(* Logix 5000 project; controller CIP vendor 1 type 14 code 106 rev 20.12; software revision 20.06; part 12 of 13 *)
(* tags used below, declared in another part *)
   Alarm_Present : INT[8];
   Bit : BOOL[128];
   Counter : COUNTER[10];
   Level_Bits : BOOL[32];
   Level_Timers : TIMER[20];
   MOA_OFF : DINT[10];
   MOA_ON : DINT[10];
   MOA_ONS : DINT;
   MOA_Screen1_Auto : BOOL;
   MOA_Screen1_Man_Off : BOOL;
   MOA_Screen1_Man_On : BOOL;
   MOA_Screen2_Auto : BOOL;
   MOA_Screen2_Man_Off : BOOL;
   MOA_Screen2_Man_On : BOOL;
   MOA_Screen3_Auto : BOOL;
   MOA_Screen3_Man_Off : BOOL;
   MOA_Screen3_Man_On : BOOL;
   MOA_Screen4_Auto : BOOL;
   MOA_Screen4_Man_Off : BOOL;
   MOA_Screen4_Man_On : BOOL;
   MOA_Select : DINT[10];
   MOA_Status : DINT[10];
   MOA_Temp : DINT;
   OpCode_Pin : DINT[5];
   Panelview : INT[40];
   Recipe : RECIPE[41];
   SCLD_Drain_PH : REAL;
   SCLD_Dryer_Duct_Temp : REAL;
   SCLD_Dryer_Exhaust_Temp : REAL;
   SCLD_Return_Temp : REAL;
   SCLD_Rinse_Cond : REAL;
   SCLD_Solution_Tank_Lvl : REAL;
   SCLD_Supply_Temp : REAL;
   SCLD_Wash_Cond : REAL;
   SP_Dryer_Min_Temp : REAL;
   SP_Dryer_Temp : REAL;
   SP_Return_Temp : REAL;
   SP_Rinse_Cond : REAL;
   SP_Solution_Tank_Fill_Lvl : REAL;
   SP_Solution_Tank_Lvl : REAL;
   SP_Supply_Temp : REAL;
   SP_Wash_Cond : REAL;
   SP_Wash_Cond_Hold : REAL;
   Timer : TIMER[99];
   Utility_Out : DINT[5];
   WashChamberDoorGasketCTRL : DINT;
(* MainProgram, continued *)

ROUTINE _30_MAN_OFF_AUTO   (* ladder *)
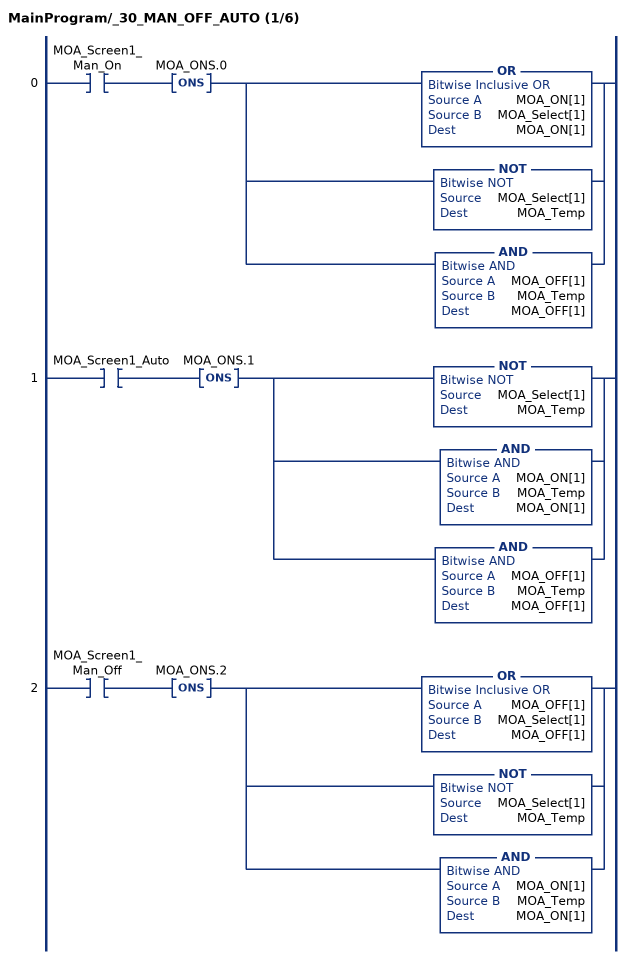
   0: XIC(MOA_Screen1_Man_On)ONS(MOA_ONS.0)[OR(MOA_ON[1],MOA_Select[1],MOA_ON[1]) ,NOT(MOA_Select[1],MOA_Temp) ,AND(MOA_OFF[1],MOA_Temp,MOA_OFF[1]) ];
   1: XIC(MOA_Screen1_Auto)ONS(MOA_ONS.1)[NOT(MOA_Select[1],MOA_Temp) ,AND(MOA_ON[1],MOA_Temp,MOA_ON[1]) ,AND(MOA_OFF[1],MOA_Temp,MOA_OFF[1]) ];
   2: XIC(MOA_Screen1_Man_Off)ONS(MOA_ONS.2)[OR(MOA_OFF[1],MOA_Select[1],MOA_OFF[1]) ,NOT(MOA_Select[1],MOA_Temp) ,AND(MOA_ON[1],MOA_Temp,MOA_ON[1]) ];
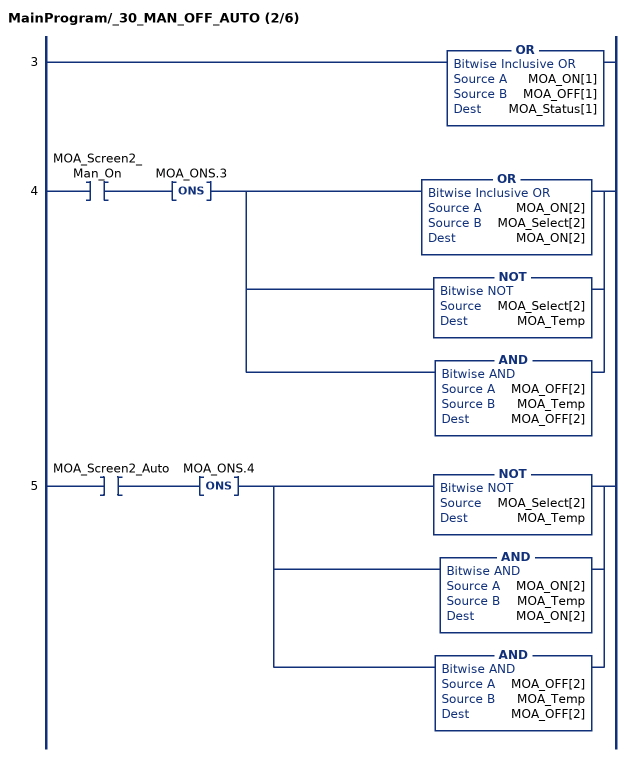
   3: OR(MOA_ON[1],MOA_OFF[1],MOA_Status[1]);
   4: XIC(MOA_Screen2_Man_On)ONS(MOA_ONS.3)[OR(MOA_ON[2],MOA_Select[2],MOA_ON[2]) ,NOT(MOA_Select[2],MOA_Temp) ,AND(MOA_OFF[2],MOA_Temp,MOA_OFF[2]) ];
   5: XIC(MOA_Screen2_Auto)ONS(MOA_ONS.4)[NOT(MOA_Select[2],MOA_Temp) ,AND(MOA_ON[2],MOA_Temp,MOA_ON[2]) ,AND(MOA_OFF[2],MOA_Temp,MOA_OFF[2]) ];
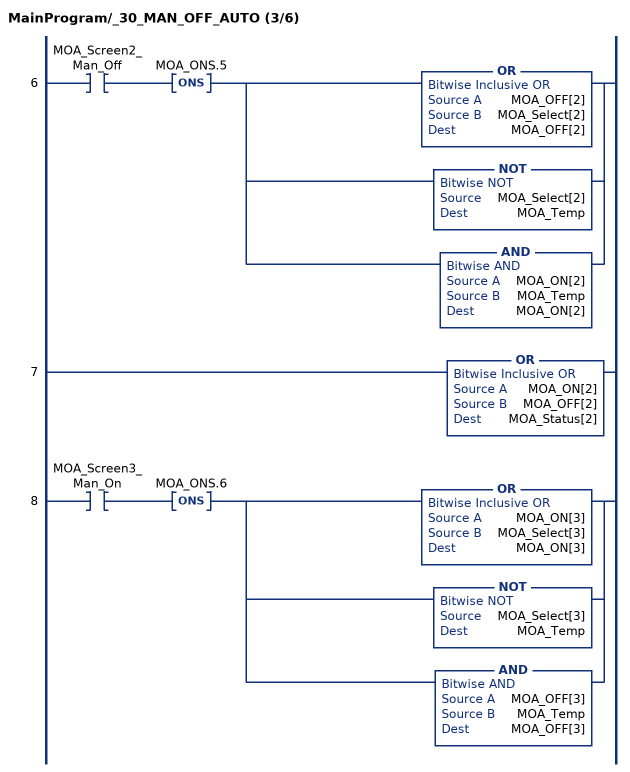
   6: XIC(MOA_Screen2_Man_Off)ONS(MOA_ONS.5)[OR(MOA_OFF[2],MOA_Select[2],MOA_OFF[2]) ,NOT(MOA_Select[2],MOA_Temp) ,AND(MOA_ON[2],MOA_Temp,MOA_ON[2]) ];
   7: OR(MOA_ON[2],MOA_OFF[2],MOA_Status[2]);
   8: XIC(MOA_Screen3_Man_On)ONS(MOA_ONS.6)[OR(MOA_ON[3],MOA_Select[3],MOA_ON[3]) ,NOT(MOA_Select[3],MOA_Temp) ,AND(MOA_OFF[3],MOA_Temp,MOA_OFF[3]) ];
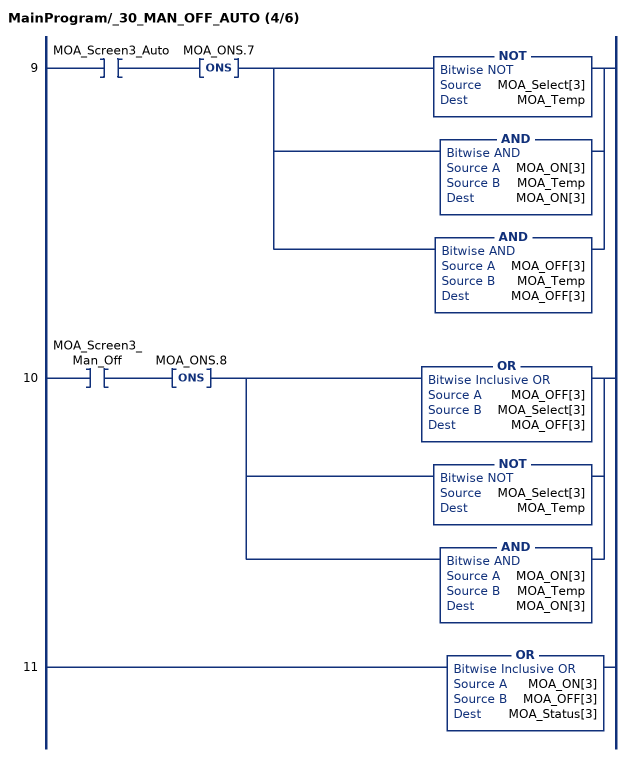
   9: XIC(MOA_Screen3_Auto)ONS(MOA_ONS.7)[NOT(MOA_Select[3],MOA_Temp) ,AND(MOA_ON[3],MOA_Temp,MOA_ON[3]) ,AND(MOA_OFF[3],MOA_Temp,MOA_OFF[3]) ];
   10: XIC(MOA_Screen3_Man_Off)ONS(MOA_ONS.8)[OR(MOA_OFF[3],MOA_Select[3],MOA_OFF[3]) ,NOT(MOA_Select[3],MOA_Temp) ,AND(MOA_ON[3],MOA_Temp,MOA_ON[3]) ];
   11: OR(MOA_ON[3],MOA_OFF[3],MOA_Status[3]);
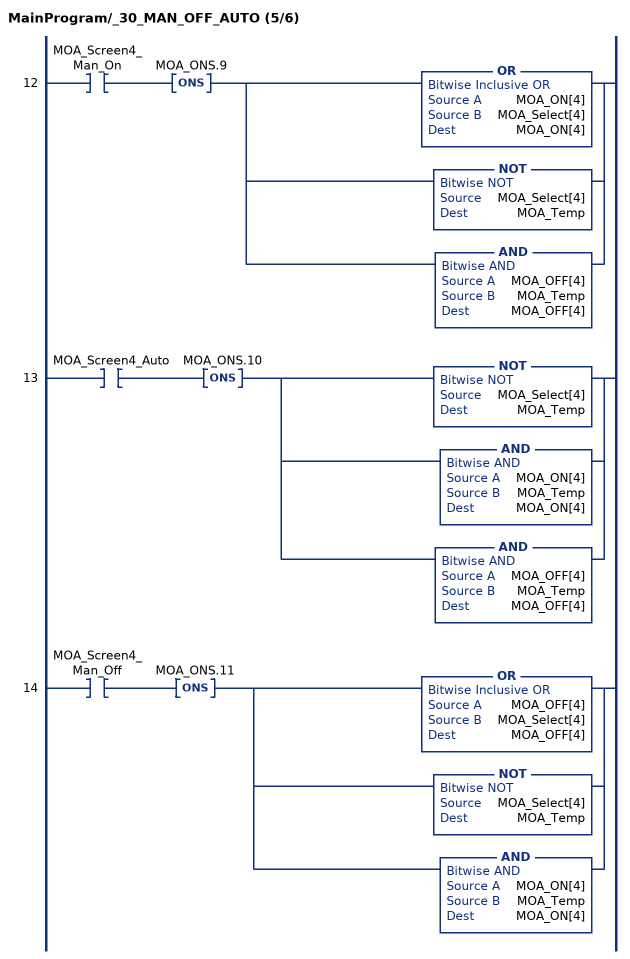
   12: XIC(MOA_Screen4_Man_On)ONS(MOA_ONS.9)[OR(MOA_ON[4],MOA_Select[4],MOA_ON[4]) ,NOT(MOA_Select[4],MOA_Temp) ,AND(MOA_OFF[4],MOA_Temp,MOA_OFF[4]) ];
   13: XIC(MOA_Screen4_Auto)ONS(MOA_ONS.10)[NOT(MOA_Select[4],MOA_Temp) ,AND(MOA_ON[4],MOA_Temp,MOA_ON[4]) ,AND(MOA_OFF[4],MOA_Temp,MOA_OFF[4]) ];
   14: XIC(MOA_Screen4_Man_Off)ONS(MOA_ONS.11)[OR(MOA_OFF[4],MOA_Select[4],MOA_OFF[4]) ,NOT(MOA_Select[4],MOA_Temp) ,AND(MOA_ON[4],MOA_Temp,MOA_ON[4]) ];
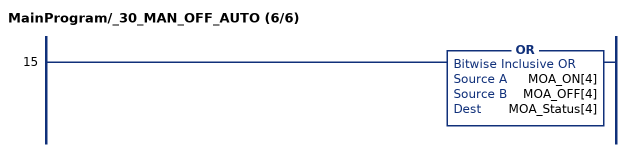
   15: OR(MOA_ON[4],MOA_OFF[4],MOA_Status[4]);
END_ROUTINE

ROUTINE _80_DOOR_GASKET   (* ladder *)
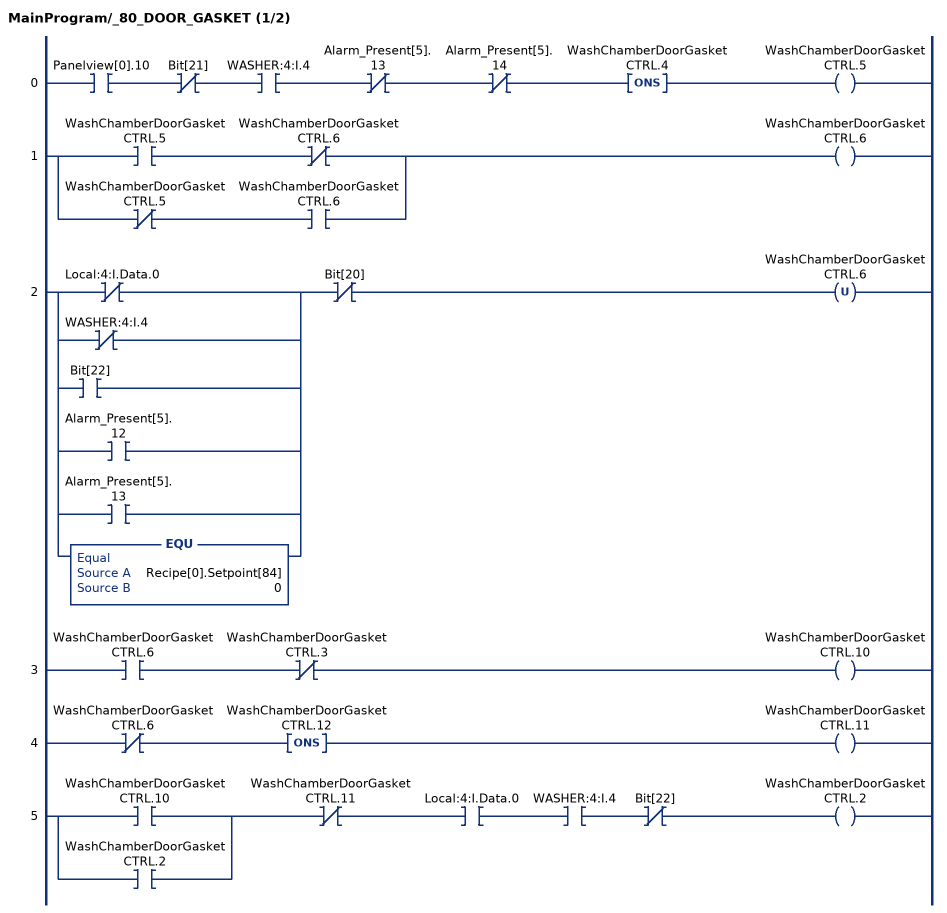
   0: XIC(Panelview[0].10)XIO(Bit[21])XIC(WASHER:4:I.4)XIO(Alarm_Present[5].13)XIO(Alarm_Present[5].14)ONS(WashChamberDoorGasketCTRL.4)OTE(WashChamberDoorGasketCTRL.5);
   1: [XIC(WashChamberDoorGasketCTRL.5) XIO(WashChamberDoorGasketCTRL.6) ,XIO(WashChamberDoorGasketCTRL.5) XIC(WashChamberDoorGasketCTRL.6) ]OTE(WashChamberDoorGasketCTRL.6);
   2: [XIO(Local:4:I.Data.0) ,XIO(WASHER:4:I.4) ,XIC(Bit[22]) ,XIC(Alarm_Present[5].12) ,XIC(Alarm_Present[5].13) ,EQU(Recipe[0].Setpoint[84],0) ]XIO(Bit[20])OTU(WashChamberDoorGasketCTRL.6);
   3: XIC(WashChamberDoorGasketCTRL.6)XIO(WashChamberDoorGasketCTRL.3)OTE(WashChamberDoorGasketCTRL.10);
   4: XIO(WashChamberDoorGasketCTRL.6)ONS(WashChamberDoorGasketCTRL.12)OTE(WashChamberDoorGasketCTRL.11);
   5: [XIC(WashChamberDoorGasketCTRL.10) ,XIC(WashChamberDoorGasketCTRL.2) ]XIO(WashChamberDoorGasketCTRL.11)XIC(Local:4:I.Data.0)XIC(WASHER:4:I.4)XIO(Bit[22])OTE(WashChamberDoorGasketCTRL.2);
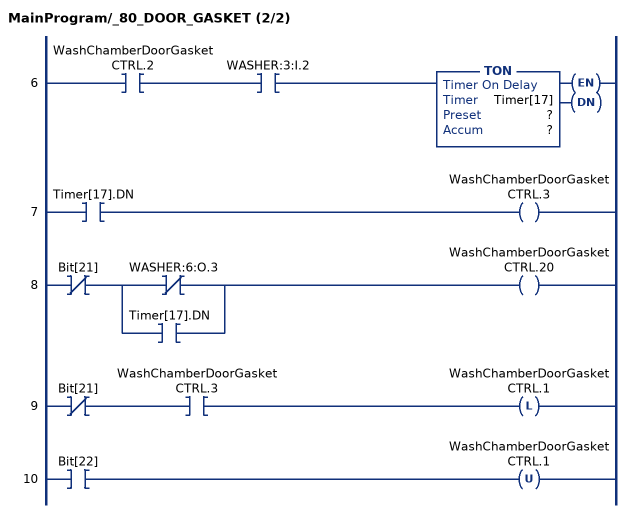
   6: XIC(WashChamberDoorGasketCTRL.2)XIC(WASHER:3:I.2)TON(Timer[17],?,?);
   7: XIC(Timer[17].DN)OTE(WashChamberDoorGasketCTRL.3);
   8: XIO(Bit[21])[XIO(WASHER:6:O.3) ,XIC(Timer[17].DN) ]OTE(WashChamberDoorGasketCTRL.20);
   9: XIO(Bit[21])XIC(WashChamberDoorGasketCTRL.3)OTL(WashChamberDoorGasketCTRL.1);
   10: XIC(Bit[22])OTU(WashChamberDoorGasketCTRL.1);
END_ROUTINE

ROUTINE _86_TEMPERATURE   (* ladder *)
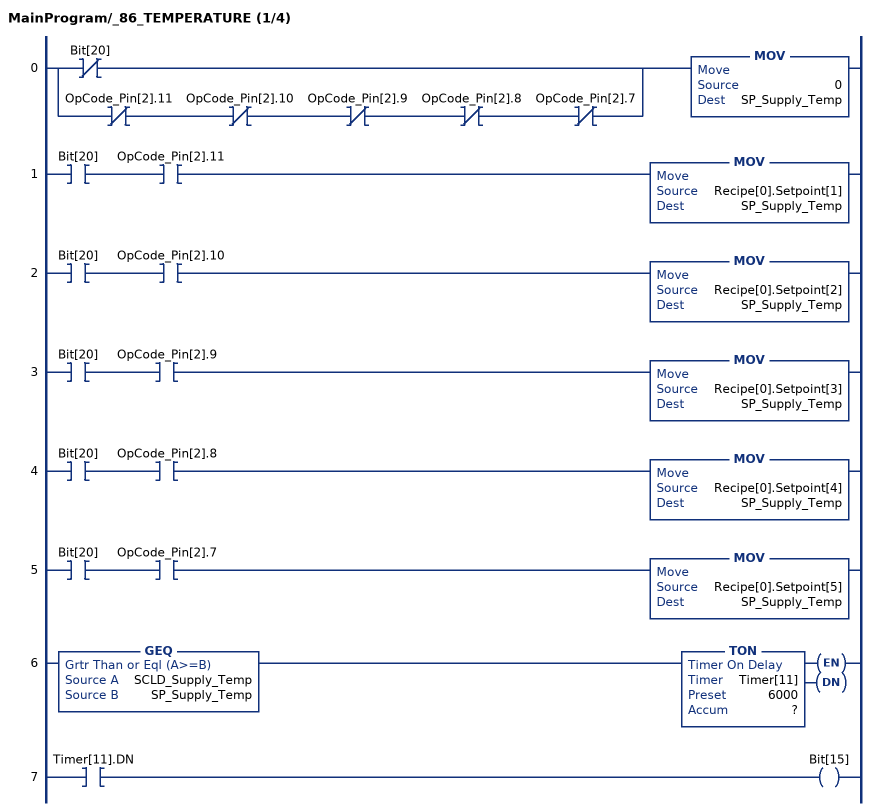
   0: [XIO(Bit[20]) ,XIO(OpCode_Pin[2].11) XIO(OpCode_Pin[2].10) XIO(OpCode_Pin[2].9) XIO(OpCode_Pin[2].8) XIO(OpCode_Pin[2].7) ]MOV(0,SP_Supply_Temp);
   1: XIC(Bit[20])XIC(OpCode_Pin[2].11)MOV(Recipe[0].Setpoint[1],SP_Supply_Temp);
   2: XIC(Bit[20])XIC(OpCode_Pin[2].10)MOV(Recipe[0].Setpoint[2],SP_Supply_Temp);
   3: XIC(Bit[20])XIC(OpCode_Pin[2].9)MOV(Recipe[0].Setpoint[3],SP_Supply_Temp);
   4: XIC(Bit[20])XIC(OpCode_Pin[2].8)MOV(Recipe[0].Setpoint[4],SP_Supply_Temp);
   5: XIC(Bit[20])XIC(OpCode_Pin[2].7)MOV(Recipe[0].Setpoint[5],SP_Supply_Temp);
   6: GEQ(SCLD_Supply_Temp,SP_Supply_Temp)TON(Timer[11],?,?);
   7: XIC(Timer[11].DN)OTE(Bit[15]);
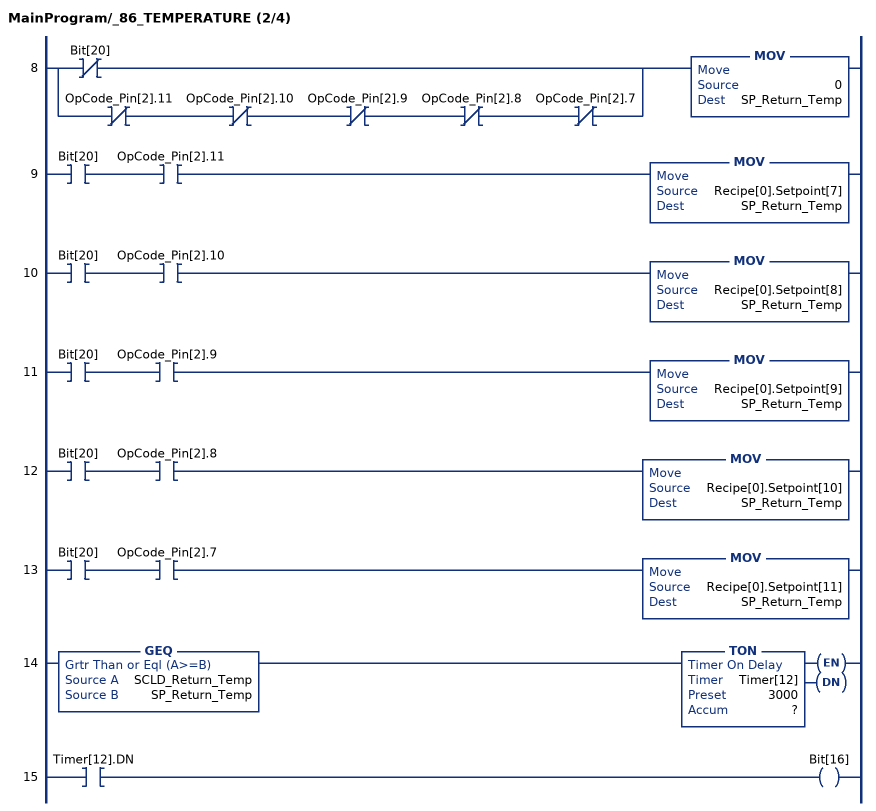
   8: [XIO(Bit[20]) ,XIO(OpCode_Pin[2].11) XIO(OpCode_Pin[2].10) XIO(OpCode_Pin[2].9) XIO(OpCode_Pin[2].8) XIO(OpCode_Pin[2].7) ]MOV(0,SP_Return_Temp);
   9: XIC(Bit[20])XIC(OpCode_Pin[2].11)MOV(Recipe[0].Setpoint[7],SP_Return_Temp);
   10: XIC(Bit[20])XIC(OpCode_Pin[2].10)MOV(Recipe[0].Setpoint[8],SP_Return_Temp);
   11: XIC(Bit[20])XIC(OpCode_Pin[2].9)MOV(Recipe[0].Setpoint[9],SP_Return_Temp);
   12: XIC(Bit[20])XIC(OpCode_Pin[2].8)MOV(Recipe[0].Setpoint[10],SP_Return_Temp);
   13: XIC(Bit[20])XIC(OpCode_Pin[2].7)MOV(Recipe[0].Setpoint[11],SP_Return_Temp);
   14: GEQ(SCLD_Return_Temp,SP_Return_Temp)TON(Timer[12],?,?);
   15: XIC(Timer[12].DN)OTE(Bit[16]);
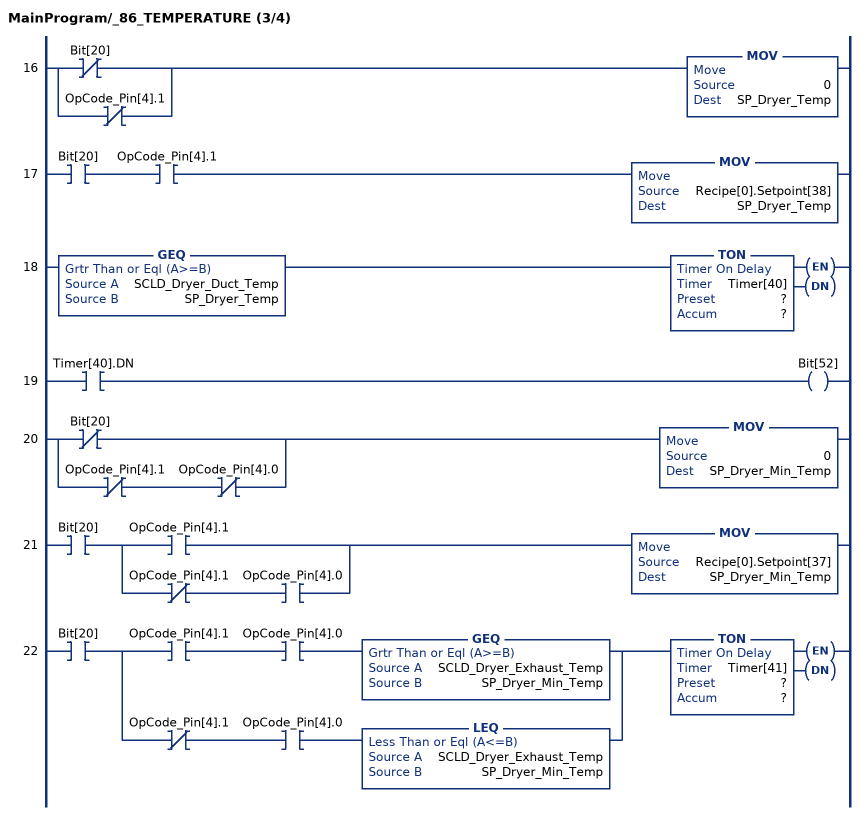
   16: [XIO(Bit[20]) ,XIO(OpCode_Pin[4].1) ]MOV(0,SP_Dryer_Temp);
   17: XIC(Bit[20])XIC(OpCode_Pin[4].1)MOV(Recipe[0].Setpoint[38],SP_Dryer_Temp);
   18: GEQ(SCLD_Dryer_Duct_Temp,SP_Dryer_Temp)TON(Timer[40],?,?);
   19: XIC(Timer[40].DN)OTE(Bit[52]);
   20: [XIO(Bit[20]) ,XIO(OpCode_Pin[4].1) XIO(OpCode_Pin[4].0) ]MOV(0,SP_Dryer_Min_Temp);
   21: XIC(Bit[20])[XIC(OpCode_Pin[4].1) ,XIO(OpCode_Pin[4].1) XIC(OpCode_Pin[4].0) ]MOV(Recipe[0].Setpoint[37],SP_Dryer_Min_Temp);
   22: XIC(Bit[20])[XIC(OpCode_Pin[4].1) XIC(OpCode_Pin[4].0) GEQ(SCLD_Dryer_Exhaust_Temp,SP_Dryer_Min_Temp) ,XIO(OpCode_Pin[4].1) XIC(OpCode_Pin[4].0) LEQ(SCLD_Dryer_Exhaust_Temp,SP_Dryer_Min_Temp) ]TON(Timer[41],?,?);
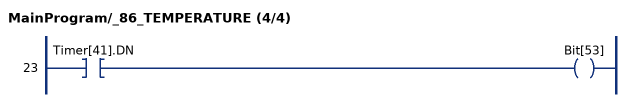
   23: XIC(Timer[41].DN)OTE(Bit[53]);
END_ROUTINE

ROUTINE _87_CONDUCTIVITY   (* ladder *)
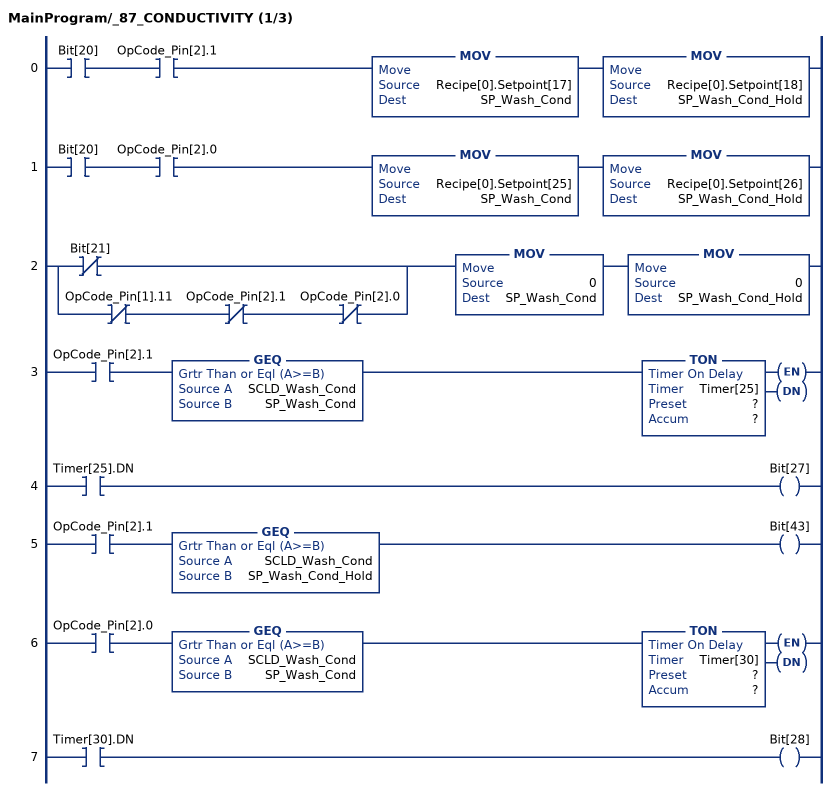
   0: XIC(Bit[20])XIC(OpCode_Pin[2].1)MOV(Recipe[0].Setpoint[17],SP_Wash_Cond)MOV(Recipe[0].Setpoint[18],SP_Wash_Cond_Hold);
   1: XIC(Bit[20])XIC(OpCode_Pin[2].0)MOV(Recipe[0].Setpoint[25],SP_Wash_Cond)MOV(Recipe[0].Setpoint[26],SP_Wash_Cond_Hold);
   2: [XIO(Bit[21]) ,XIO(OpCode_Pin[1].11) XIO(OpCode_Pin[2].1) XIO(OpCode_Pin[2].0) ]MOV(0,SP_Wash_Cond)MOV(0,SP_Wash_Cond_Hold);
   3: XIC(OpCode_Pin[2].1)GEQ(SCLD_Wash_Cond,SP_Wash_Cond)TON(Timer[25],?,?);
   4: XIC(Timer[25].DN)OTE(Bit[27]);
   5: XIC(OpCode_Pin[2].1)GEQ(SCLD_Wash_Cond,SP_Wash_Cond_Hold)OTE(Bit[43]);
   6: XIC(OpCode_Pin[2].0)GEQ(SCLD_Wash_Cond,SP_Wash_Cond)TON(Timer[30],?,?);
   7: XIC(Timer[30].DN)OTE(Bit[28]);
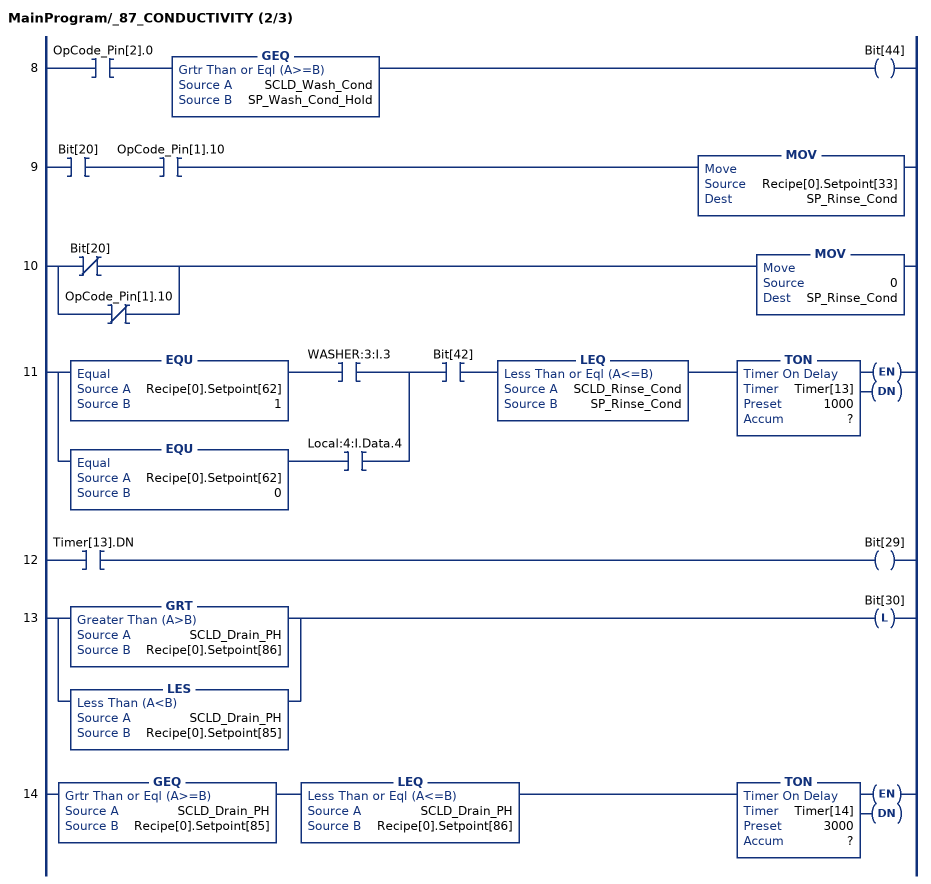
   8: XIC(OpCode_Pin[2].0)GEQ(SCLD_Wash_Cond,SP_Wash_Cond_Hold)OTE(Bit[44]);
   9: XIC(Bit[20])XIC(OpCode_Pin[1].10)MOV(Recipe[0].Setpoint[33],SP_Rinse_Cond);
   10: [XIO(Bit[20]) ,XIO(OpCode_Pin[1].10) ]MOV(0,SP_Rinse_Cond);
   11: [EQU(Recipe[0].Setpoint[62],1) XIC(WASHER:3:I.3) ,EQU(Recipe[0].Setpoint[62],0) XIC(Local:4:I.Data.4) ]XIC(Bit[42])LEQ(SCLD_Rinse_Cond,SP_Rinse_Cond)TON(Timer[13],?,?);
   12: XIC(Timer[13].DN)OTE(Bit[29]);
   13: [GRT(SCLD_Drain_PH,Recipe[0].Setpoint[86]) ,LES(SCLD_Drain_PH,Recipe[0].Setpoint[85]) ]OTL(Bit[30]);
   14: GEQ(SCLD_Drain_PH,Recipe[0].Setpoint[85])LEQ(SCLD_Drain_PH,Recipe[0].Setpoint[86])TON(Timer[14],?,?);
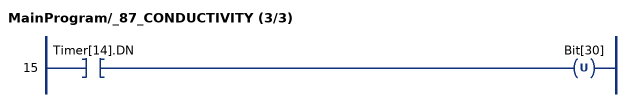
   15: XIC(Timer[14].DN)OTU(Bit[30]);
END_ROUTINE

ROUTINE _88_LEVEL   (* ladder *)
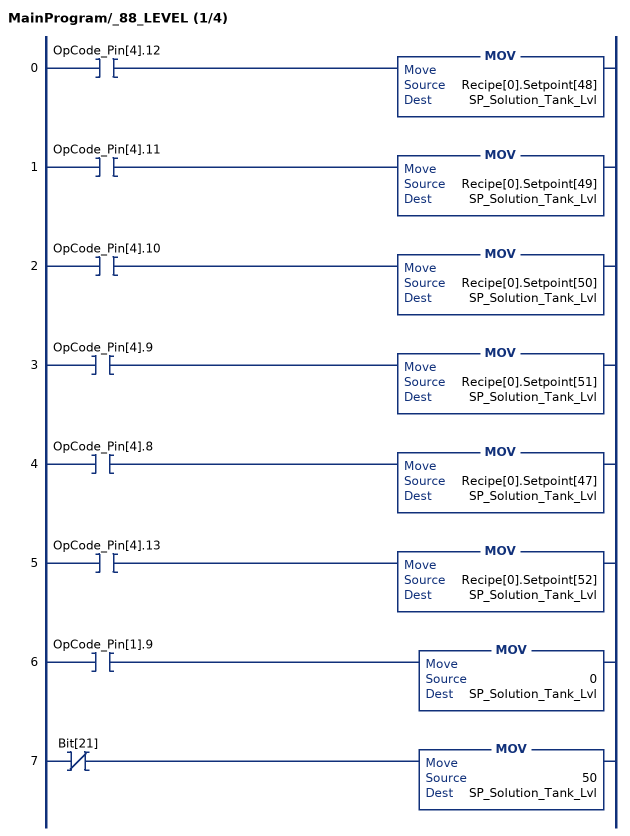
   0: XIC(OpCode_Pin[4].12)MOV(Recipe[0].Setpoint[48],SP_Solution_Tank_Lvl);
   1: XIC(OpCode_Pin[4].11)MOV(Recipe[0].Setpoint[49],SP_Solution_Tank_Lvl);
   2: XIC(OpCode_Pin[4].10)MOV(Recipe[0].Setpoint[50],SP_Solution_Tank_Lvl);
   3: XIC(OpCode_Pin[4].9)MOV(Recipe[0].Setpoint[51],SP_Solution_Tank_Lvl);
   4: XIC(OpCode_Pin[4].8)MOV(Recipe[0].Setpoint[47],SP_Solution_Tank_Lvl);
   5: XIC(OpCode_Pin[4].13)MOV(Recipe[0].Setpoint[52],SP_Solution_Tank_Lvl);
   6: XIC(OpCode_Pin[1].9)MOV(0,SP_Solution_Tank_Lvl);
   7: XIO(Bit[21])MOV(50,SP_Solution_Tank_Lvl);
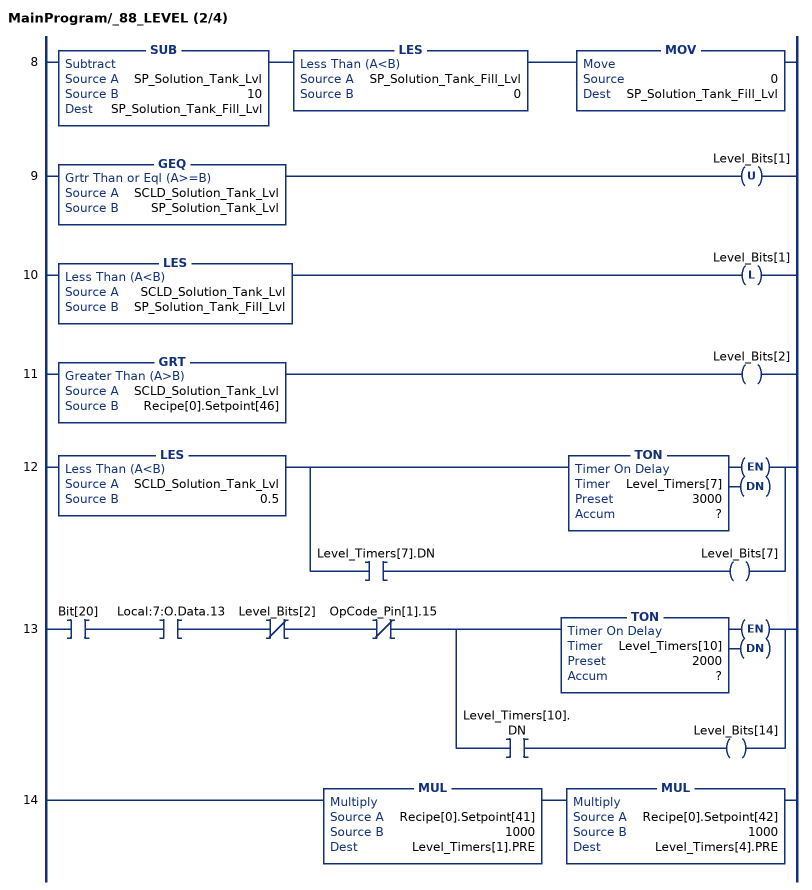
   8: SUB(SP_Solution_Tank_Lvl,10,SP_Solution_Tank_Fill_Lvl)LES(SP_Solution_Tank_Fill_Lvl,0)MOV(0,SP_Solution_Tank_Fill_Lvl);
   9: GEQ(SCLD_Solution_Tank_Lvl,SP_Solution_Tank_Lvl)OTU(Level_Bits[1]);
   10: LES(SCLD_Solution_Tank_Lvl,SP_Solution_Tank_Fill_Lvl)OTL(Level_Bits[1]);
   11: GRT(SCLD_Solution_Tank_Lvl,Recipe[0].Setpoint[46])OTE(Level_Bits[2]);
   12: LES(SCLD_Solution_Tank_Lvl,0.5)[TON(Level_Timers[7],?,?) ,XIC(Level_Timers[7].DN) OTE(Level_Bits[7]) ];
   13: XIC(Bit[20])XIC(Local:7:O.Data.13)XIO(Level_Bits[2])XIO(OpCode_Pin[1].15)[TON(Level_Timers[10],?,?) ,XIC(Level_Timers[10].DN) OTE(Level_Bits[14]) ];
   14: MUL(Recipe[0].Setpoint[41],1000,Level_Timers[1].PRE)MUL(Recipe[0].Setpoint[42],1000,Level_Timers[4].PRE);
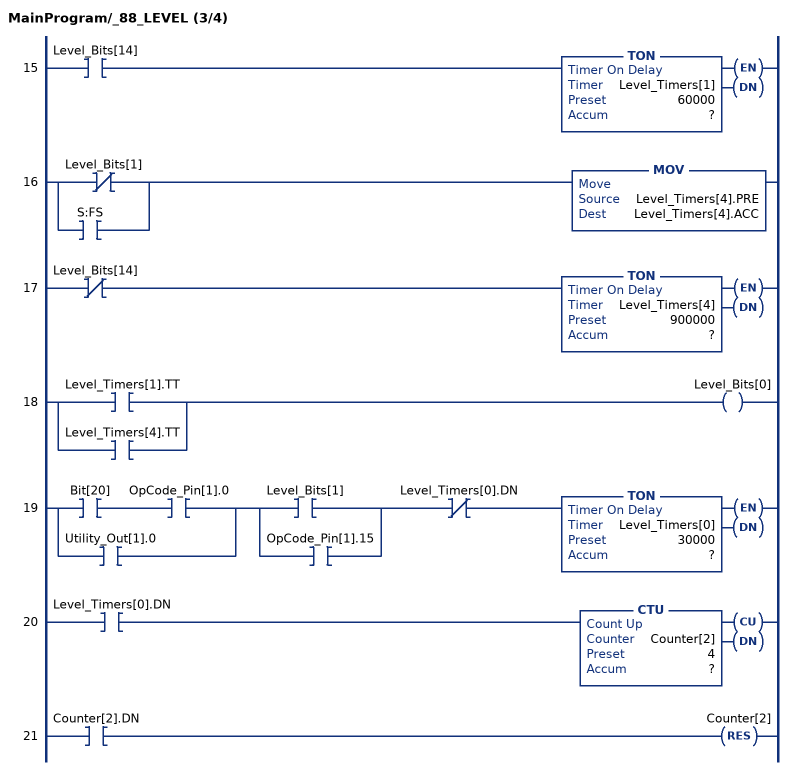
   15: XIC(Level_Bits[14])TON(Level_Timers[1],?,?);
   16: [XIO(Level_Bits[1]) ,XIC(S:FS) ]MOV(Level_Timers[4].PRE,Level_Timers[4].ACC);
   17: XIO(Level_Bits[14])TON(Level_Timers[4],?,?);
   18: [XIC(Level_Timers[1].TT) ,XIC(Level_Timers[4].TT) ]OTE(Level_Bits[0]);
   19: [XIC(Bit[20]) XIC(OpCode_Pin[1].0) ,XIC(Utility_Out[1].0) ][XIC(Level_Bits[1]) ,XIC(OpCode_Pin[1].15) ]XIO(Level_Timers[0].DN)TON(Level_Timers[0],?,?);
   20: XIC(Level_Timers[0].DN)CTU(Counter[2],?,?);
   21: XIC(Counter[2].DN)RES(Counter[2]);
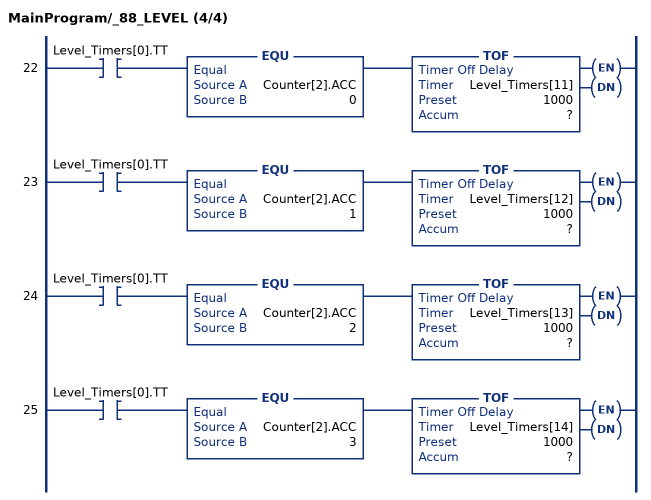
   22: XIC(Level_Timers[0].TT)EQU(Counter[2].ACC,0)TOF(Level_Timers[11],?,?);
   23: XIC(Level_Timers[0].TT)EQU(Counter[2].ACC,1)TOF(Level_Timers[12],?,?);
   24: XIC(Level_Timers[0].TT)EQU(Counter[2].ACC,2)TOF(Level_Timers[13],?,?);
   25: XIC(Level_Timers[0].TT)EQU(Counter[2].ACC,3)TOF(Level_Timers[14],?,?);
END_ROUTINE
